(*
SPDX-FileCopyrightText: © 2026 Oleksandr Tiutyk <trofimich@gmail.com>
SPDX-License-Identifier: MIT
License: https://opensource.org/license/mit
*)

(*!
<summary>Identifies the execution lifecycle of a test element.</summary>
*)

{attribute 'qualified_only'}
{attribute 'strict'}
{attribute 'to_string'}
TYPE TEST_ELEMENT_STATE :
(
	READY,
	RUNNING,
	COMPLETED
);
END_TYPE

(* stored: Version 1.1.0.1
   DUT TEST_ELEMENT_STATE: Id {a458aadb-286f-44a1-910a-0030333bba25} *)
